// TIA Portal V20 export
// export: Created 2026-10-19T18:45:46.61206Z, ExportSetting None, DisplayName Totally Integrated Automation Portal, DisplayVersion V20 Update 6, DisplayName TIA Portal Openness, DisplayVersion V20 Update 6, DisplayName TIA Portal Version Control Interface, DisplayVersion V20 Update 6, DisplayName SINAMICS Startdrive Advanced, DisplayVersion V20 SP1, DisplayName SINAMICS Startdrive G130, G150, S120, S150, SINAMICS MV, G220, S200, S210, DisplayVersion V20 SP1, DisplayName SINAMICS Startdrive G110M, G120, G120C, G120D, G120P, G115D, DisplayVersion V20 SP1, DisplayName STEP 7 Professional, DisplayVersion V20 Update 6, DisplayName STEP 7 Safety, DisplayVersion V20 Update 2, DisplayName WinCC Basic/Comfort/Advanced, DisplayVersion V20 Update 6, DisplayName WinCC Unified, DisplayVersion V20 Update 6
VAR_GLOBAL   // PLC tag table "IO_Charger Panel_L2"
   "CHARGER L2 - Output Voltage" AT %ID788 : Real;   // Actual Output Voltage
   "CHARGER L2 - Output Current" AT %ID792 : Real;   // Actual Output Current
   "CHARGER L2 - Set Voltage Feedback" AT %ID796 : Real;   // Set Voltage Value
   "CHARGER L2 - Set Current Feedback" AT %ID800 : Real;   // Set Current Value
   "CHARGER L2 - Charging Start" AT %I804.0 : Bool;   // Charging Running Status
   "CHARGER L2 - Set Voltage Output" AT %QD292 : Real;   // Issue Target Voltage
   "CHARGER L2 - Set Current Output" AT %QD296 : Real;   // Issue Target Current
   "CHARGER L2 - Start Charging" AT %Q300.0 : Bool;   // Start Charging Command
   "CHARGER L2 - Stop Charging" AT %Q300.1 : Bool;   // Stop Charging Command
   "CHARGER L2 - Confirm Voltage & Current Setting" AT %Q300.2 : Bool;   // Confirmation Command
END_VAR
